Fanuc KAREL source: KT00164.KL

PROGRAM KT00164
%NOLOCKGROUP
VAR
  I1: INTEGER
  R2: REAL
  OUT: REAL
BEGIN
  I1 = 2
    R2 = 3.0
  OUT = I1 MOD R2
END KT00164
